SUBAPPLICATION Uebung_161 (* Übung zu logiBUS_ENC_ID: Inkrementalgeber zählen, Taster setzt zurück *)
  (* Standard: 61499-2; Description: Copyright (c) 2026 Meisterschulen am Ostbahnhof This program and the accompanying materials are made available under the terms of the Eclipse Public License 2.0 which is available at https://www.eclipse.org/legal/epl-2.0/ SPDX-License-Identifier: EPL-2.0 *)
  (* Version 1.0, 2026-11-26, Franz Höpfinger, Meisterschulen am Ostbahnhof, initial API and implementation and/or initial documentation *)
  PACKAGE Uebungen;
  IMPORT logiBUS::io::ENC::logiBUS_ENC::Encoder_E1;
  IMPORT logiBUS::io::DI::logiBUS_DI::Input_I9;
  IMPORT logiBUS::io::DI::logiBUS_DI_Events::BUTTON_SINGLE_CLICK;
  IMPORT logiBUS::io::DQ::logiBUS_DO::Output_Q1;
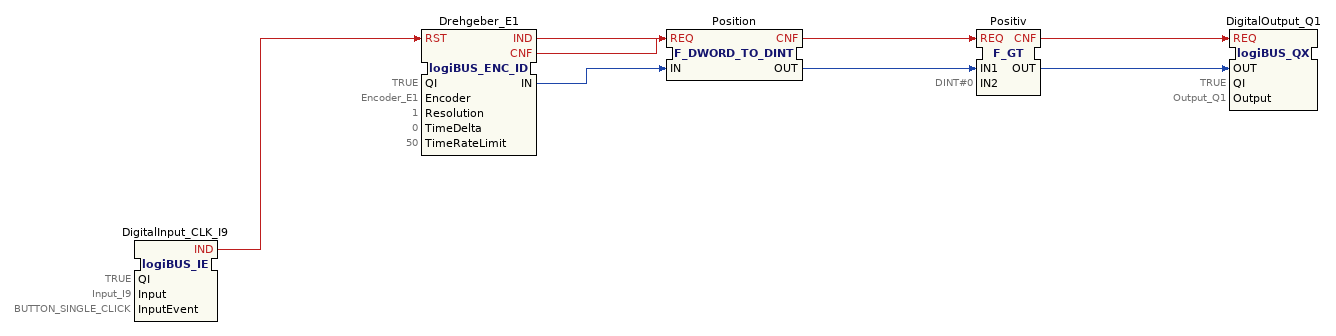
  (* Inkrementalgeber (logiBUS_ENC_ID) am Trainer20: A = GPIO22, B = GPIO23, Taster = I9. Drehen: IND mit der Position in IN (DWORD). F_DWORD_TO_DINT macht daraus die vorzeichenbehaftete Position (Watch: Position.OUT). Q1 an = Position größer 0. I9 Klick: RST setzt die Position auf 0. Resolution 1 = ein Schritt je Raste, 2 oder 4 = feiner. TimeRateLimit 50 ms: höchstens ein IND je 50 ms. Andere Boards melden STATUS 'this board has no encoder E1'. *)
  FBS
    Drehgeber_E1 : logiBUS::io::ENC::logiBUS_ENC_ID(QI := TRUE, Encoder := Encoder_E1, Resolution := 1, TimeDelta := 0, TimeRateLimit := 50); (* Trainer20: A = GPIO22, B = GPIO23 *)
    Position : iec61131::conversion::F_DWORD_TO_DINT; (* IN (DWORD) als vorzeichenbehaftete Position *)
    Positiv : iec61131::comparison::F_GT(IN2 := DINT#0); (* Position größer 0? *)
    DigitalOutput_Q1 : logiBUS::io::DQ::logiBUS_QX(QI := TRUE, Output := Output_Q1); (* an = Position größer 0 *)
    DigitalInput_CLK_I9 : logiBUS::io::DI::logiBUS_IE(QI := TRUE, Input := Input_I9, InputEvent := BUTTON_SINGLE_CLICK); (* Taster am Drehgeber (GPIO24) *)
  END_FBS
  EVENT_CONNECTIONS
    Drehgeber_E1.IND TO Position.REQ;
    Drehgeber_E1.CNF TO Position.REQ;
    Position.CNF TO Positiv.REQ;
    Positiv.CNF TO DigitalOutput_Q1.REQ;
    DigitalInput_CLK_I9.IND TO Drehgeber_E1.RST;
  END_CONNECTIONS
  DATA_CONNECTIONS
    Drehgeber_E1.IN TO Position.IN;
    Position.OUT TO Positiv.IN1;
    Positiv.OUT TO DigitalOutput_Q1.OUT;
  END_CONNECTIONS
END_SUBAPPLICATION
